Fanuc KAREL source: KT00821.KL

PROGRAM KT00821
%NOLOCKGROUP
VAR
  I1: INTEGER
  I2: INTEGER
  OUT: REAL
BEGIN
  I1 = 2
  I2 = 3
  I1 = 2
  I2 = 3
  OUT = SIN(I1)
END KT00821
